Fanuc KAREL source: KD00011.KL

PROGRAM KD00011
%NOLOCKGROUP
VAR
  I: INTEGER
  J: INTEGER
  B: BOOLEAN
  R: REAL
  S: STRING[80]
BEGIN
  ATTACH
END KD00011
